Fanuc KAREL source: KA00173.KL

PROGRAM KA00173
%NOLOCKGROUP
VAR
  SRC: ARRAY[4] OF STRING[20]
  DST: ARRAY[4] OF REAL
BEGIN
  DST = SRC
END KA00173
